FUNCTION_BLOCK FB_NCICimasa_SampleBox EXTENDS FB_RecipeBase

METHOD Build : BOOL
VAR
END_VAR
VAR_INST
    nBuildStep : INT;
    machineConfig : ST_GantryXYZ_Config;
    
    // Zmienne do obsługi kopiowania
    fbFileCopy : FB_FileCopy;
    sUsbPath   : STRING(255) := '\Hard Disk2\vrg_flash\Cimasa_SampleBox.nc';
    sPlcPath   : STRING(255) := '\Hard Disk\GCode\Cimasa_SampleBox.nc';
END_VAR
Build := FALSE;

CASE nBuildStep OF
    0:
        _Busy := TRUE;
        _Done := FALSE;
        _Error := FALSE;
        
        // Rozpoczęcie kopiowania z pendrive'a (Hard Disk2) na dysk PLC
        fbFileCopy(
            sSrcPathName  := sUsbPath,
            sDestPathName := sPlcPath,
            bExecute      := TRUE
        );
        
        nBuildStep := 10;

    10:
        fbFileCopy(bExecute := FALSE); // Opuszczenie flagi Execute
        
        // Oczekiwanie na zakończenie pracy bloku kopiującego
        IF NOT fbFileCopy.bBusy THEN
            IF fbFileCopy.bError THEN
                // Błąd kopiowania (np. brak USB lub pliku) - logujemy i idziemy dalej
                ADSLOGSTR(ADSLOG_MSGTYPE_WARN, 'No flash.', '');
            ELSE
                // Sukces - plik został nadpisany nową wersją z USB
                ADSLOGSTR(ADSLOG_MSGTYPE_HINT, 'NCno  flash.', '');
            END_IF
            
            // Niezależnie od wyniku (błąd czy sukces), recepta wskazuje na plik lokalny
            _Config.GCodePath := sPlcPath; 
            
            nBuildStep := 1000;
        END_IF

    1000:
        _Busy := FALSE;
        _Done := TRUE; 
        nBuildStep := 0;
        Build := TRUE;
        
END_CASE
END_METHOD

PROPERTY ExecutionRoute : E_ExecutionRoute
GET
ExecutionRoute := E_ExecutionRoute.eGCode;
END_GET
END_PROPERTY

END_FUNCTION_BLOCK

(* stored: Version 1.1.0.1, ProductVersion 3.1.4024.15
   POU FB_NCICimasa_SampleBox: Id {e495bbc6-186b-41e3-b55e-5390c6a836f8}, SpecialFunc None
   Method Build: Id {aa1e595f-ced9-4a60-89fc-140c3e1dd111}
   Property ExecutionRoute: Id {6a4eba19-6c0e-4358-a0ad-58b76747b17e}
   Get Get: Id {d7d2ba43-db8b-4ed8-951b-8e6102f5a71e} *)
